TYPE TcoKukaKssPn_IO_v_9_3_x :
STRUCT
	PnIoBoxState AT %I*	:	UINT;
	PnIoBoxDiag AT %I*	:	UINT;
	PnIoBoxCtrl AT %Q*	:	UINT;
	{attribute addProperty Name "<#IN#>"}
	In : TcoKukaKss_Inputs_v_9_3_x;
	{attribute addProperty Name "<#OUT#>"}
	Out : TcoKukaKss_Outputs_v_9_3_x;
END_STRUCT
END_TYPE

(* stored: Version 1.1.0.1, ProductVersion 3.1.4024.12
   DUT TcoKukaKssPn_IO_v_9_3_x: Id {7d2ee15a-b7ae-493a-9504-6a2004a42de5} *)
